{attribute 'qualified_only'}
{attribute 'strict'}
{attribute 'to_string'}
TYPE E_ActuatorModulatingFunctionParam : // Use for passing parameters into modulating actuator functions
(
	None		:= 0, //unused
	Position	:= 1 //target position in %
);
END_TYPE

(* stored: Version 1.1.0.1, ProductVersion 3.1.4024.12
   DUT E_ActuatorModulatingFunctionParam: Id {de60f522-0e11-4f61-aa71-feeb2d5b52dd} *)
